(* PLC project Vn_networks2_edit_swapped, Beckhoff Automation GmbH TwinCAT PLC Control 3.5.13.21 *)
(* stored: creationDateTime 1970-01-01T00:00:00 *)

PROGRAM Vn_networks2_edit_swapped

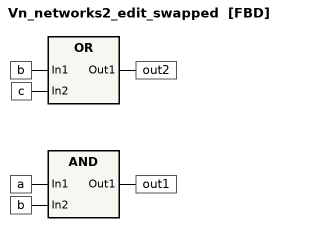
(* FBD diagram, written out as Structured Text *)
out2 := b OR c;
out1 := a AND b;
END_PROGRAM
